FUNCTION_BLOCK FB_BatchSteps (* Migrated from IEC 61131-3 ST *)
  (* Standard: 61499-2 *)
  (* Version 1.0, 2026-11-06, st2fb *)
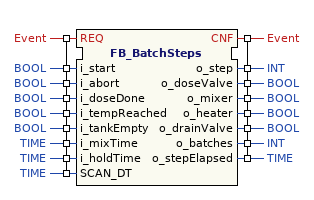
  EVENT_INPUT
    REQ WITH i_start, i_abort, i_doseDone, i_tempReached, i_tankEmpty, i_mixTime, i_holdTime, SCAN_DT;
  END_EVENT
  EVENT_OUTPUT
    CNF WITH o_step, o_doseValve, o_mixer, o_heater, o_drainValve, o_batches, o_stepElapsed;
  END_EVENT
  VAR_INPUT
    i_start : BOOL;
    i_abort : BOOL;
    i_doseDone : BOOL;
    i_tempReached : BOOL;
    i_tankEmpty : BOOL;
    i_mixTime : TIME;
    i_holdTime : TIME;
    SCAN_DT : TIME;
  END_VAR
  VAR_OUTPUT
    o_step : INT;
    o_doseValve : BOOL;
    o_mixer : BOOL;
    o_heater : BOOL;
    o_drainValve : BOOL;
    o_batches : INT;
    o_stepElapsed : TIME;
  END_VAR
  VAR
    ST2FB_NOW : TIME := T#0s;
    statStepTimer_IN : BOOL := FALSE;
    statStepTimer_PT : TIME := T#0s;
    statStepTimer_Q : BOOL := FALSE;
    statStepTimer_ET : TIME := T#0s;
    statStepTimer_STATE : INT := 0;
    statStepTimer_PREV_IN : BOOL := FALSE;
    statStepTimer_START_TIME : TIME := T#0s;
    statBatchCounter_CU : BOOL := FALSE;
    statBatchCounter_R : BOOL := FALSE;
    statBatchCounter_PV : INT := 0;
    statBatchCounter_Q : BOOL := FALSE;
    statBatchCounter_CV : INT := 0;
    statBatchCounter_CU_T_Q : BOOL := FALSE;
    statBatchCounter_CU_T_M : BOOL := FALSE;
    statStartEdge_CLK : BOOL := FALSE;
    statStartEdge_Q : BOOL := FALSE;
    statStartEdge_M : BOOL := FALSE;
    statStepTimerRun : BOOL := FALSE;
    statBatchDone : BOOL := FALSE;
    statStepPreset : TIME := T#0s;
  END_VAR
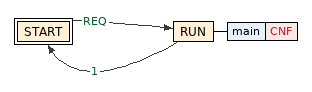
  EC_STATES
    START;
    RUN : main -> CNF;
  END_STATES
  EC_TRANSITIONS
    START TO RUN := REQ;
    RUN TO START := 1;
  END_TRANSITIONS
  ALGORITHM main IN ST:
ST2FB_NOW := ST2FB_NOW + SCAN_DT;

statStartEdge_CLK := i_start;
statStartEdge_Q := statStartEdge_CLK AND NOT statStartEdge_M;
statStartEdge_M := statStartEdge_CLK;

statStepTimer_IN := statStepTimerRun;
statStepTimer_PT := statStepPreset;
IF (statStepTimer_STATE = 0) AND NOT statStepTimer_PREV_IN AND statStepTimer_IN THEN
  statStepTimer_STATE := 1;
  statStepTimer_Q := FALSE;
  statStepTimer_START_TIME := ST2FB_NOW;
ELSE
  IF NOT statStepTimer_IN THEN
    statStepTimer_ET := T#0s;
    statStepTimer_Q := FALSE;
    statStepTimer_STATE := 0;
  ELSIF statStepTimer_STATE = 1 THEN
    IF statStepTimer_START_TIME + statStepTimer_PT <= ST2FB_NOW THEN
      statStepTimer_STATE := 2;
      statStepTimer_Q := TRUE;
      statStepTimer_ET := statStepTimer_PT;
    ELSE
      statStepTimer_ET := ST2FB_NOW - statStepTimer_START_TIME;
    END_IF;
  END_IF;
END_IF;
statStepTimer_PREV_IN := statStepTimer_IN;
o_stepElapsed := statStepTimer_ET;

o_doseValve := FALSE;
o_mixer := FALSE;
o_heater := FALSE;
o_drainValve := FALSE;
statBatchDone := FALSE;
IF i_abort AND o_step <> 0 THEN
  o_step := 90;
  statStepTimerRun := FALSE;
END_IF;

CASE o_step OF
  0:
    IF statStartEdge_Q AND NOT i_abort THEN
      o_step := 10;
    END_IF;
  10:
    o_doseValve := TRUE;
    IF i_doseDone THEN
      o_step := 20;
      statStepPreset := i_mixTime;
      statStepTimerRun := TRUE;
    END_IF;
  20:
    o_mixer := TRUE;
    IF statStepTimer_Q THEN
      statStepTimerRun := FALSE;
      o_step := 30;
    END_IF;
  30:
    o_mixer := TRUE;
    o_heater := TRUE;
    IF i_tempReached THEN
      o_step := 40;
      statStepPreset := i_holdTime;
      statStepTimerRun := TRUE;
    END_IF;
  40:
    o_mixer := TRUE;
    o_heater := NOT i_tempReached;
    IF statStepTimer_Q THEN
      statStepTimerRun := FALSE;
      o_step := 50;
    END_IF;
  50:
    o_drainValve := TRUE;
    IF i_tankEmpty THEN
      statBatchDone := TRUE;
      o_step := 0;
    END_IF;
  90:
    o_drainValve := TRUE;
    IF i_tankEmpty AND NOT i_abort THEN
      o_step := 0;
    END_IF;
ELSE
  o_step := 0;
END_CASE;

statBatchCounter_CU := statBatchDone;
statBatchCounter_R := FALSE;
statBatchCounter_PV := 500;
statBatchCounter_CU_T_Q := statBatchCounter_CU AND NOT statBatchCounter_CU_T_M;
statBatchCounter_CU_T_M := statBatchCounter_CU;
IF statBatchCounter_R THEN
  statBatchCounter_CV := 0;
ELSIF statBatchCounter_CU_T_Q AND (statBatchCounter_CV < statBatchCounter_PV) THEN
  statBatchCounter_CV := statBatchCounter_CV + 1;
END_IF;
statBatchCounter_Q := statBatchCounter_CV >= statBatchCounter_PV;
o_batches := statBatchCounter_CV;
  END_ALGORITHM
END_FUNCTION_BLOCK
